Fanuc KAREL source: kt00090.KL

-- PROVISIONAL review KL for V770-1; original PC SHA256 5449f94839e0ccee222e246b7a210cd059eaf5f4c26544682d079a6874965722
-- Incomplete behavior may be omitted. Consult companion uncertainty JSON. Do not deploy.
PROGRAM KT00090
%NOLOCKGROUP
VAR
  I2 : INTEGER
  OUT : REAL
-- UNRESOLVED_DECL H1 type=002017
BEGIN
  -- UNRESOLVED_PC offsets 5-19; opcodes 2E,22,9D,33,B4
  -- UNRESOLVED_PC offsets 24-35; opcodes 2E,23
  -- UNRESOLVED_PC offsets 40-63; opcodes 22,9D,33,B3,21,54,64,23
  -- UNRESOLVED_PC offsets 68-72; opcodes 7F
END KT00090
